(* IEC 61131-3 sources: Lasal-MCP/examples/SampleSource/LASALScreenAdvancedSolution/LASALScreenAdvancedSolution/LASALScreenAdvacnedSolution/Stations/Terminal/HMI/Class/IconSourceList, 1 file *)

(* ---- IconSourceList.st ---- *)
(*!
<Class
	Name               = "IconSourceList"
	Revision           = "0.0"
	RealtimeTask       = "false"
	CyclicTask         = "false"
	BackgroundTask     = "false"
	Sigmatek           = "false"
	OSInterface        = "false"
	HighPriority       = "false"
	Automatic          = "false"
	UpdateMode         = "Prescan"
	SharedCommandTable = "true"
	Objectsize         = "(544,120)">
	<Channels>
		<Client Name="_Grafix" Required="false" Internal="false"/>
		<Client Name="DestList" Required="true" Internal="false"/>
		<Client Name="DragDropArea" Required="true" Internal="false"/>
		<Client Name="SigCLib" Required="false" Internal="false"/>
	</Channels>
	<Network Name="IconSourceList">
		<!-- List of Components in this network -->
		<Components>
			<Object
				Name       = "_base"
				Class      = "_ScrollArea2"
				Position   = "(218,120)"
				Visualized = "true"
				Remotely   = "true">
				<Channels>
					<Server Name="ActPos"/>
					<Server Name="Refresh"/>
					<Server Name="Server0"/>
					<Client Name="ExtendedScrollBar" Value="0"/>
					<Client Name="LineHighness"/>
					<Client Name="LineWidth"/>
					<Client Name="Lse"/>
					<Client Name="VerticalLevel"/>
				</Channels>
			</Object>
		</Components>
		<Comments>
		</Comments>
		<!-- List of Connections in this network -->
		<Connections>
			<Connection Source="this.Server0" Destination="_base.Server0" Vertices="(886,210),(714,210),"/>
			<Connection Source="this.Refresh" Destination="_base.Refresh" Vertices="(886,270),(714,270),"/>
			<Connection Source="this.ActPos" Destination="_base.ActPos" Vertices="(886,330),(714,330),"/>
			<Connection Source="_base.Lse" Destination="this.Lse" Vertices="(218,210),(38,210),"/>
			<Connection Source="_base.VerticalLevel" Destination="this.VerticalLevel" Vertices="(218,270),(38,270),"/>
			<Connection Source="_base.LineWidth" Destination="this.LineWidth" Vertices="(218,330),(38,330),"/>
		</Connections>
		<!-- Headerfiles -->
		<Options>
		</Options>
	</Network>
</Class>
*)
#pragma using _ScrollArea2

IconSourceList : CLASS
: _ScrollArea2
  //Servers:
  //Clients:
	DestList 	: CltChCmd_IconDestList;
	DragDropArea 	: CltChCmd_DragDropArea;
	_Grafix 	: CltChCmd__Grafix;
	SigCLib 	: CltChCmd_SigCLib;
  //Variables:
		BackgroundColor 	: _COLOR;
		TextColor 	: _COLOR;
		FrameColor 	: _COLOR;
		IconSelected 	: BOOL;
		SelectedLineNo 	: DINT;
		SchemeNo 	: UDINT;
		myRoom 	: _ROOM;
		LastEvent 	: _EVENT;
		pImage 	: ^_BMP;
		pDragDropPio 	: ^_IO;
		pLSEpio 	: ^_IO;
		pDestListScroll 	: ^_SCROLL;
  //Functions:

	FUNCTION VIRTUAL GLOBAL Init;
				//! <Function Comment="[#ENGLISH]&#13;&#10;this method is called everytime when the input is active and a event occured&#13;&#10;&#13;&#10;ped ....... pointer to _EDITOR information&#13;&#10;pe ........ pointer to _EVENT information&#13;&#10;&#13;&#10;for the returnstatement there are 3 different possibilities&#13;&#10;_IDLE ..... the system should goon like it is (system goes on)&#13;&#10;_IDIDIT ... i did it (system is ready)&#13;&#10;_IFAILED .. i tried to do my best, but i failed (system is ready)&#13;&#10;" Name="GetEvent"/>
	FUNCTION __CDECL VIRTUAL GLOBAL GetEvent
		VAR_INPUT
			ped 	: ^_EDITOR;			//! <Variable Comment="pointer to _EDITOR information" Name="GetEvent.ped"/>
			pe 	: ^_EVENT;			//! <Variable Comment="pointer to _EVENT information" Name="GetEvent.pe"/>
		END_VAR
		VAR_OUTPUT
			retcode (EAX) 	: _DOIT;			//! <Variable Comment="for the returnstatement there are 3 different possibilities&#13;&#10;  _IDLE ..... the system should goon like it is (system goes on)&#13;&#10;  _IDIDIT ... i did it (system is ready)&#13;&#10;  _IFAILED .. i tried to do my best, but i failed (system is ready)&#13;&#10;" Name="GetEvent.retcode"/>
		END_VAR;
				//! <Function Comment="[#ENGLISH]&#13;&#10;method is called cyclic during object is on screen&#13;&#10;&#13;&#10;pio ....... pointer to io information&#13;&#10;input .... TRUE it&apos;s an input / FALSE it&apos;s an output&#13;&#10;" Name="IF_Run"/>
	FUNCTION __CDECL VIRTUAL GLOBAL IF_Run
		VAR_INPUT
			pio 	: ^_IO;			//! <Variable Comment="pointer to _IO information given by LSE" Name="IF_Run.pio"/>
			input 	: BOOL;			//! <Variable Comment="TRUE it&apos;s an input&#13;&#10;FALSE it&apos;s an output" Name="IF_Run.input"/>
		END_VAR;
				//! <Function Comment="method is called every time when redraw of a single line is necessary.&#13;&#10;" Name="Line"/>
	FUNCTION __CDECL VIRTUAL GLOBAL Line
		VAR_INPUT
			ps 	: ^_SCROLL;			//! <Variable Comment="pointer to structure _SCROLL" Name="Line.ps"/>
			pr 	: ^_ROOM;			//! <Variable Comment="pointer to place where line should be drawn" Name="Line.pr"/>
			line 	: UINT;			//! <Variable Comment="16 bit linenumber " Name="Line.line"/>
			state 	: BOOL;			//! <Variable Comment="line is selected (true) or passive (false)" Name="Line.state"/>
		END_VAR;
  //Tables:
	FUNCTION @STD
		VAR_OUTPUT
			ret_code	: CONFSTATES;
		END_VAR;
	FUNCTION GLOBAL TAB @CT_;
END_CLASS;

#pragma usingLtd _Grafix
#pragma usingLtd DragDropArea
#pragma usingLtd IconDestList
#pragma usingLtd SigCLib

FUNCTION VIRTUAL GLOBAL IconSourceList::Init

  if (_FirstScan = TRUE) then

    Scroll.position.no := 10; // nummber of lines
    Scroll.line_height := 75; // height of the line

    // colors for text, frame and background
    TextColor       := _Grafix.MakeColor(backcolor:= INVISIBLE,
                                         frontcolor:= BLACK);

    FrameColor      := _Grafix.MakeColor(backcolor:= INVISIBLE,
                                         frontcolor:= INVISIBLE);

    BackgroundColor := _Grafix.MakeColor(backcolor:= INVISIBLE,
                                         frontcolor:= INVISIBLE);
  end_if;

END_FUNCTION

FUNCTION __CDECL VIRTUAL GLOBAL IconSourceList::Line
  VAR_INPUT
		ps 	: ^_SCROLL;
		pr 	: ^_ROOM;
		line 	: UINT;
		state 	: BOOL;
	END_VAR
  VAR
  	att         :_ATTRIB;
    myImageRoom : _ROOM;
    lineNo      : ARRAY [0..10] of CHAR;
    pImage      : ^_BMP;
  END_VAR

  if (pLSEpio = NIL) then
    TRACE("pio was not assigned to pLSEpio.");
    return;
  end_if;

  if (line < Scroll.position.no) then

    _memcpy(ptr1:= #myRoom, ptr2:= ps, cntr:= sizeof(_ROOM));

    // number of the applied scheme
    SchemeNo := get_no_by_label(p0:= "DragDrop",
                                x1:= IMAGESCHEME, x2:=0);

    if (SchemeNo = DEFSCOPE) then
      TRACE("Image not found in ImageScheme 'DragDrop'");
      return;
    end_if;

    pImage$^void := NewDoScheme(x0:= IMAGESCHEME,
                                x1:= line,
                                x2:= SchemeNo);

    if (pImage <> NIL) then

      myImageRoom.xy1.x := pr^.xy1.x;
      myImageRoom.xy1.y := pr^.xy1.y;
      myImageRoom.xy2.x := pr^.xy1.x + to_int(Scroll.line_height);
      myImageRoom.xy2.y := pr^.xy2.y;

      att := T_SOLID or T_COPY or T_PROP or T_LEFTBOUND;

      out_zoom_BMP(p0:= #myImageRoom,
                   p1:= pImage,
                   x2:= att);

      // insert the line no
      myImageRoom.xy1.x := pr^.xy1.x + 76;
      myImageRoom.xy1.y := pr^.xy1.y;
      myImageRoom.xy2.x := pr^.xy1.x + 76 + 20;
      myImageRoom.xy2.y := pr^.xy2.y;

      _memset(dest:= #lineNo[0], usByte:= 0, cntr:= sizeof(lineNo));

      SigCLib.IToA(val:= line, dst:= #lineNo[0], base:= 10);

      OutTextAlign(p0:= #lineNo[0],
                   x1:= 0,
                   p1:= #myImageRoom,
                   x2:= pLSEpio^.font,
                   x3:= pLSEpio^.attrib,
                   x9:= pLSEpio^.frametype,
                   x4:= TextColor,
                   x5:= FrameColor,
                   x6:= BackgroundColor,
                   x7:= 1);
    else
      TRACE("Image not found in ImageScheme 'DragDrop'");
      return;
    end_if;

  end_if;

END_FUNCTION

FUNCTION __CDECL VIRTUAL GLOBAL IconSourceList::GetEvent
	VAR_INPUT
		ped 	: ^_EDITOR;
		pe 	: ^_EVENT;
	END_VAR
	VAR_OUTPUT
		retcode (EAX) 	: _DOIT;
	END_VAR

  pDragDropPio := DragDropArea.GetDimension();
  pDestListScroll := DestList.GetDimensionDestScroll();

  case pe^.ftype of
    //===========================================================================
    _EVENT_HIDPRESS:

      // IconSourceList icons-area
      if ((pe^.dot.x >= myRoom.xy1.x) &
          (pe^.dot.x <= myRoom.xy2.x - LEVELBUTTON_WIDTH) &
          (pe^.dot.y >= myRoom.xy1.y) &
          (pe^.dot.y <= myRoom.xy2.y)) then

        SelectedLineNo := (((pe^.dot.y - ped^.input.io.room.xy1.y)
                            / Scroll.line_height) + Scroll.position.begin);

        DragDropArea.SetLineNo(SelectedLine:= SelectedLineNo);
        // selected icon
        DragDropArea.SetIcon(SelectedLine:= SelectedLineNo);
        IconSelected := TRUE;

      // IconSourceList Scroll-Area
      elsif ((pe^.dot.x >= myRoom.xy2.x - LEVELBUTTON_WIDTH) &
             (pe^.dot.x <= myRoom.xy2.x) &
             (pe^.dot.y >= myRoom.xy1.y) &
             (pe^.dot.y <= myRoom.xy2.y)) then

        // stop drawing
        DragDropArea.DeleteIcon();
        IconSelected := FALSE;

        Refresh := 1;
        retcode := _IDIDIT;
      end_if;

    //===========================================================================
    _EVENT_HIDMOVE:

      _memcpy(ptr1:= #lastEvent,
              ptr2:= pe,
              cntr:= sizeof(lastEvent));

      // draw icon
      if (IconSelected = TRUE) then

        DragDropArea.DrawIcon(CoordX:= pe^.dot.x,
                              CoordY:= pe^.dot.y);
      end_if;

    //===========================================================================
    _EVENT_HIDRELEASE:
      // IconDestList icon-area
      if ((lastEvent.dot.x >= pDestListScroll^.out_room.xy1.x) &
          (lastEvent.dot.x <= pDestListScroll^.out_room.xy2.x - LEVELBUTTON_WIDTH) &
          (lastEvent.dot.y >= pDestListScroll^.out_room.xy1.y) &
          (lastEvent.dot.y <= pDestListScroll^.out_room.xy2.y)) then

         DestList.InsertIcon(IconNo:= SelectedLineNo,
                             pEvent:= #lastEvent);
      end_if;

      // stop drawing
      DragDropArea.ClearScreen();
      DragDropArea.DeleteIcon();
      IconSelected := FALSE;

      Refresh := 1;
      retcode := _IDIDIT;

  end_case;

  // call base class
  retcode := _ScrollArea2::GetEvent(ped:= ped, pe:= pe);

END_FUNCTION

FUNCTION __CDECL VIRTUAL GLOBAL IconSourceList::IF_Run
	VAR_INPUT
		pio 	: ^_IO;
		input 	: BOOL;
	END_VAR

  pLSEpio := pio;

  _ScrollArea2::IF_Run(pio:= pio, input:= input);

END_FUNCTION
